(* IEC 61131-3 sources: Test-Git_ESME26/TestProgettoESME_26.fbsproj/AxisModuleLib Migration/LibraryDiagnostics, 1 file *)

(* ---- AXM_FC_EtDiagExtToString.fn.st ---- *)
FUNCTION AXM_FC_EtDiagExtToString : STRING[80]
VAR_INPUT
	i_etDiagExt : AXM_ET_DiagExt;
END_VAR
VAR_OUTPUT
	q_etDiag	: GD.ET_Diag := GD.ET_Diag.Ok;
	q_etDiagExt	: AXM_ET_DiagExt := AXM_ET_DiagExt.Ok;
END_VAR
VAR
END_VAR

AXM_FC_EtDiagExtToString := TO_STRING(i_etDiagExt);
IF TO_UDINT(AXM_FC_EtDiagExtToString) <> 0 THEN // if the string is not a number the result is 0
	AXM_FC_EtDiagExtToString := Standard.CONCAT('Unknown DiagExt: ', TO_STRING(i_etDiagExt));
	q_etDiag := GD.ET_Diag.InputParameterInvalid;
	q_etDiagExt := AXM_ET_DiagExt.DiagExtRange;
END_IF
